(* IEC 61131-3 sources: llm-plc-st-eval/data/processed_definitivo/gemini-3.1-pro-preview/A2/zero_shot, 3 files *)

(* ---- ejec_1.st ---- *)
FUNCTION_BLOCK FB_Batch
VAR_INPUT
    nivelA : BOOL;
    nivelB : BOOL;
    nivelVacio : BOOL;
    btnInicio : BOOL;
    btnAbort : BOOL;
    temp : REAL;
END_VAR

VAR_OUTPUT
    vA : BOOL;
    vB : BOOL;
    calentador : BOOL;
    mezclador : BOOL;
    vDescarga : BOOL;
    fase : INT := 0;
END_VAR

VAR
    timerMezcla : TON;
    trigInicio : R_TRIG;
    trigAbort : R_TRIG;
END_VAR

// Detección de flancos para los botones
trigInicio(CLK := btnInicio);
trigAbort(CLK := btnAbort);

// Lógica de Aborto (ignorado en reposo, fase = 0)
IF trigAbort.Q AND fase > 0 THEN
    IF NOT nivelVacio THEN
        fase := 5; // Pasa a descarga si hay producto en el reactor
    ELSE
        fase := 0; // Vuelve a reposo directo si ya está vacío
    END_IF;
END_IF;

// Máquina de estados secuencial
CASE fase OF
    0: // Fase 0: Reposo
        IF trigInicio.Q THEN
            fase := 1;
        END_IF;

    1: // Fase 1: Dosificar componente A
        IF nivelA THEN
            fase := 2;
        END_IF;

    2: // Fase 2: Dosificar componente B
        IF nivelB THEN
            fase := 3;
        END_IF;

    3: // Fase 3: Calentar
        IF temp >= 60.0 THEN
            fase := 4;
        END_IF;

    4: // Fase 4: Mezclar
        IF timerMezcla.Q THEN
            fase := 5;
        END_IF;

    5: // Fase 5: Descargar
        IF nivelVacio THEN
            fase := 0;
        END_IF;
END_CASE;

// Temporizador de mezcla (se activa únicamente durante la fase 4)
timerMezcla(IN := (fase = 4), PT := T#120S);

// Asignación de salidas (se cierran/apagan automáticamente al cambiar de fase)
vA := (fase = 1);
vB := (fase = 2);
calentador := (fase = 3);
mezclador := (fase = 4);
vDescarga := (fase = 5);

END_FUNCTION_BLOCK

(* ---- ejec_2.st ---- *)
FUNCTION_BLOCK FB_Batch
VAR_INPUT
    nivelA : BOOL;      (* Sensor de nivel del componente A *)
    nivelB : BOOL;      (* Sensor de nivel del componente B *)
    nivelVacio : BOOL;  (* Sensor de reactor vacío *)
    btnInicio : BOOL;   (* Botón para iniciar la receta *)
    btnAbort : BOOL;    (* Botón para abortar la receta *)
    temp : REAL;        (* Temperatura actual del reactor *)
END_VAR

VAR_OUTPUT
    vA : BOOL;          (* Válvula del componente A *)
    vB : BOOL;          (* Válvula del componente B *)
    calentador : BOOL;  (* Actuador del calentador *)
    mezclador : BOOL;   (* Actuador del mezclador *)
    vDescarga : BOOL;   (* Válvula de descarga *)
    fase : INT := 0;    (* Fase actual de la receta (0 a 5) *)
END_VAR

VAR
    timerMezcla : TON;  (* Temporizador para la fase de mezcla *)
END_VAR

(* Actualización del temporizador: se activa solo durante la fase 4 *)
timerMezcla(IN := (fase = 4), PT := T#120S);

(* Lógica de Aborto: activa en cualquier fase de 1 a 5 *)
IF btnAbort AND (fase >= 1) AND (fase <= 5) THEN
    IF NOT nivelVacio THEN
        fase := 5; (* Si hay producto, pasa a descargar *)
    ELSE
        fase := 0; (* Si ya está vacío, pasa a reposo directo *)
    END_IF;
END_IF;

(* Máquina de estados de la receta secuencial *)
CASE fase OF
    0: (* Fase 0: Reposo *)
        IF btnInicio THEN
            fase := 1;
        END_IF;

    1: (* Fase 1: Dosificar A *)
        IF nivelA THEN
            fase := 2;
        END_IF;

    2: (* Fase 2: Dosificar B *)
        IF nivelB THEN
            fase := 3;
        END_IF;

    3: (* Fase 3: Calentar *)
        IF temp >= 60.0 THEN
            fase := 4;
        END_IF;

    4: (* Fase 4: Mezclar *)
        IF timerMezcla.Q THEN
            fase := 5;
        END_IF;

    5: (* Fase 5: Descargar *)
        IF nivelVacio THEN
            fase := 0;
        END_IF;
ELSE
    (* Estado seguro en caso de valor fuera de rango *)
    fase := 0;
END_CASE;

(* Control de salidas físicas basado en la fase activa *)
(* Al evaluar al final, un aborto cierra las válvulas y actuadores de inmediato *)
vA := (fase = 1);
vB := (fase = 2);
calentador := (fase = 3);
mezclador := (fase = 4);
vDescarga := (fase = 5);

END_FUNCTION_BLOCK

(* ---- ejec_3.st ---- *)
FUNCTION_BLOCK FB_Batch
VAR_INPUT
    nivelA     : BOOL; // Sensor de nivel alcanzado para componente A
    nivelB     : BOOL; // Sensor de nivel alcanzado para componente B
    nivelVacio : BOOL; // Sensor de reactor vacío
    btnInicio  : BOOL; // Botón para iniciar la receta
    btnAbort   : BOOL; // Botón para abortar el proceso
    temp       : REAL; // Temperatura actual del reactor
END_VAR

VAR_OUTPUT
    vA         : BOOL; // Válvula de dosificación componente A
    vB         : BOOL; // Válvula de dosificación componente B
    calentador : BOOL; // Actuador del calentador
    mezclador  : BOOL; // Actuador del mezclador
    vDescarga  : BOOL; // Válvula de descarga
    fase       : INT;  // Fase actual del proceso (0 a 5)
END_VAR

VAR
    TON_Mezcla : TON;  // Temporizador para la fase de mezclado
END_VAR

// ---------------------------------------------------------
// Lógica de Aborto
// ---------------------------------------------------------
IF btnAbort AND fase > 0 THEN
    IF fase <> 5 THEN
        IF NOT nivelVacio THEN
            fase := 5; // Si hay producto, pasar a descarga
        ELSE
            fase := 0; // Si está vacío, pasar a reposo
        END_IF;
    END_IF;
    // Si la fase ya es 5, el aborto no hace nada y continúa la descarga
END_IF;

// ---------------------------------------------------------
// Máquina de Estados (Receta)
// ---------------------------------------------------------
CASE fase OF
    0: // Fase 0: Reposo
        IF btnInicio THEN
            fase := 1;
        END_IF;

    1: // Fase 1: Dosificar componente A
        IF nivelA THEN
            fase := 2;
        END_IF;

    2: // Fase 2: Dosificar componente B
        IF nivelB THEN
            fase := 3;
        END_IF;

    3: // Fase 3: Calentar
        IF temp >= 60.0 THEN
            fase := 4;
        END_IF;

    4: // Fase 4: Mezclar
        IF TON_Mezcla.Q THEN
            fase := 5;
        END_IF;

    5: // Fase 5: Descargar
        IF nivelVacio THEN
            fase := 0;
        END_IF;
END_CASE;

// ---------------------------------------------------------
// Actualización de Temporizadores
// ---------------------------------------------------------
// El temporizador solo avanza cuando la fase activa es la 4
TON_Mezcla(IN := (fase = 4), PT := T#120S);

// ---------------------------------------------------------
// Asignación de Salidas
// ---------------------------------------------------------
// Las salidas se activan exclusivamente en su fase correspondiente.
// Un aborto cierra inmediatamente vA, vB, calentador y mezclador al cambiar la fase.
vA         := (fase = 1);
vB         := (fase = 2);
calentador := (fase = 3);
mezclador  := (fase = 4);
vDescarga  := (fase = 5);

END_FUNCTION_BLOCK
